// ============================================================================
// DB_1001_MachineMode_DJ005.scl - FB_1001_MachineMode_BufferFraming_DJ005 的背景数据块 (V15.1.0, 2026-11-15)
// ============================================================================
// 功能说明: 模式 / 暂停 / 停止 / 机器级报警。
//   背景 DB 不写变量, 变量来自 FB; 由 OB1 调用 "DB_1001_MachineMode_DJ005"(...) 时使用。
//   TIA 全局 DB 里不能放 FB 实例, 故每个功能块一个背景 DB (LSP-905 §4.11)。
// ============================================================================

DATA_BLOCK "DB_1001_MachineMode_DJ005"
"FB_1001_MachineMode_BufferFraming_DJ005"
BEGIN
END_DATA_BLOCK
